(* IEC 61131-3 sources: bcs-engineering-dsl/language/test/generating/edge_detection_test/expected, 2 files *)

(* ---- MAIN_decl.st ---- *)
PROGRAM MAIN
VAR
    TestEdgeDetection_sensor1: BOOL;
    TestEdgeDetection_sensor2: BOOL;
    TestEdgeDetection_pushButton: BOOL;
    TestEdgeDetection_startSignal: BOOL;
    TestEdgeDetection_stopSignal: BOOL;
    TestEdgeDetection_toggleOutput: BOOL;
    TestEdgeDetection_pulseOutput: BOOL := FALSE;
    R_TRIG_Instance1: R_TRIG;
    F_TRIG_Instance2: F_TRIG;
    R_TRIG_Instance3: R_TRIG;
    R_TRIG_Instance4: R_TRIG;
    F_TRIG_Instance5: F_TRIG;
END_VAR

(* ---- MAIN_impl.st ---- *)
// Control Unit 'TestEdgeDetection'
R_TRIG_Instance1(CLK := TestEdgeDetection_sensor1);
IF R_TRIG_Instance1.Q THEN
    TestEdgeDetection_startSignal := TRUE;
END_IF;
F_TRIG_Instance2(CLK := TestEdgeDetection_sensor2);
IF F_TRIG_Instance2.Q THEN
    TestEdgeDetection_stopSignal := TRUE;
END_IF;
R_TRIG_Instance3(CLK := TestEdgeDetection_pushButton);
IF R_TRIG_Instance3.Q THEN
    TestEdgeDetection_toggleOutput := NOT TestEdgeDetection_toggleOutput;
END_IF;
R_TRIG_Instance4(CLK := TestEdgeDetection_sensor1);
IF R_TRIG_Instance4.Q THEN
    TestEdgeDetection_pulseOutput := TRUE;
END_IF;
F_TRIG_Instance5(CLK := TestEdgeDetection_sensor2);
IF F_TRIG_Instance5.Q THEN
    TestEdgeDetection_pulseOutput := TRUE;
END_IF;
